(*
	Samples every span, as the OpenTelemetry AlwaysOn sampler does, even the child of a parent
	that was not sampled.
*)
FUNCTION_BLOCK FB_Sampler_AlwaysOn EXTENDS FB_Sampler

METHOD onStart
VAR_INPUT
	span: REFERENCE TO FB_Span;
END_VAR
span.setSampled(TRUE);
END_METHOD

END_FUNCTION_BLOCK

(* stored: Version 1.1.0.1
   POU FB_Sampler_AlwaysOn: Id {7902e1e9-d6cf-4e8b-a557-a46c357aa6c9}, SpecialFunc None
   Method onStart: Id {baf77f4c-0401-4f86-812f-9ccb21a900e3} *)
